(* IEC 61131-3 sources: vespera/src/DUT, 16 files *)

(* ---- ST_BunkerHmi.st ---- *)
(* 8 регистров, адрес = 1100 + (индекс-1)*8 *)
TYPE ST_BunkerHmi :
STRUCT
    wSts      : WORD;   (* +0 маски GVL_Const.BS_* *)
    wAlm      : WORD;   (* +1 GVL_Const.BA_SF *)
    wBypass   : WORD;   (* +2 GVL_Const.BY_DVU *)
    uTDvu     : UINT;   (* +3 с *)
    uTRestart : UINT;   (* +4 с *)
    uRes5     : UINT;
    uRes6     : UINT;
    uRes7     : UINT;
END_STRUCT
END_TYPE

(* ---- ST_BunkerIn.st ---- *)
TYPE ST_BunkerIn :
STRUCT
    xDVU : BOOL;   (* 1 = верхний уровень *)
    xDNU : BOOL;   (* 1 = продукт на нижнем уровне (для бункера поз.27 - второй датчик) *)
    xSF  : BOOL;   (* станции TORBA: 1 = автомат пульта управления включен *)
END_STRUCT
END_TYPE

(* ---- ST_BunkerPar.st ---- *)
TYPE ST_BunkerPar :
STRUCT
    wBypass   : WORD;   (* GVL_Const.BY_DVU - ДВУ отключен *)
    uTDvu     : UINT;   (* задержка срабатывания ДВУ, с *)
    uTRestart : UINT;   (* задержка повторного пуска после снятия ДВУ, с *)
END_STRUCT
END_TYPE

(* ---- ST_GlobHmi.st ---- *)
(* Общий блок, %MW0..%MW31 *)
TYPE ST_GlobHmi :
STRUCT
    wCmd        : WORD;  (* +0  маски GVL_Const.G_* *)
    wSts        : WORD;  (* +1  маски GVL_Const.GS_* *)
    wAlm        : WORD;  (* +2  аварийные стопы 1..10 (биты 0..9), 10 пожар, 11 фазы *)
    wWarn       : WORD;  (* +3  маски GVL_Const.GW_* *)
    uHeartbeat  : UINT;  (* +4  счётчик секунд, контроль связи *)
    uTPreStart  : UINT;  (* +5  предпусковой сигнал, с *)
    uTDksGrace  : UINT;  (* +6  разгон до контроля ДКС, с *)
    uTDksPulse  : UINT;  (* +7  нет импульсов ДКС, 0.1 с *)
    uTFcFb      : UINT;  (* +8  нет сигнала работы ПЧ, с *)
    uTFsStart   : UINT;  (* +9  нет статуса фотосепаратора после пуска, с *)
    uTGateMove  : UINT;  (* +10 контроль хода заслонки поз.1, с *)
    uSirenOn    : UINT;  (* +11 1 = аварийная сирена разрешена *)
    uRes        : ARRAY[12..31] OF UINT;
END_STRUCT
END_TYPE

(* ---- ST_GlobPar.st ---- *)
TYPE ST_GlobPar :
STRUCT
    uTPreStart : UINT;
    uTDksGrace : UINT;
    uTDksPulse : UINT;   (* 0.1 с *)
    uTFcFb     : UINT;
    uTFsStart  : UINT;
    uTGateMove : UINT;
    uSirenOn   : UINT;
END_STRUCT
END_TYPE

(* ---- ST_Link.st ---- *)
(* Связь "механизм подаёт на ..." для блокировок и последовательностей *)
TYPE ST_Link :
STRUCT
    iFrom    : INT;    (* индекс механизма-источника *)
    eTo      : INT;    (* GVL_Const.LT_MECH / LT_BUNKER / LT_INVALID *)
    iTo      : INT;    (* индекс механизма или бункера *)
    xProduct : BOOL;   (* TRUE - поток продукта (пауза по ДВУ распространяется назад),
                          FALSE - вспомогательная связь (аспирация, отходы) *)
END_STRUCT
END_TYPE

(* ---- ST_MechCfg.st ---- *)
(* Постоянная конфигурация механизма *)
TYPE ST_MechCfg :
STRUCT
    eKind     : INT;     (* GVL_Const.K_DOL / K_FC / K_GATE / K_FS *)
    xHasQF    : BOOL;    (* контроль автомата защиты (QF/SF) *)
    eDks      : INT;     (* GVL_Const.DKS_NONE / DKS_PULSE / DKS_LEVEL *)
    xHasDSL   : BOOL;    (* датчики сбегания ленты 1 и 2 *)
    xHasDP    : BOOL;    (* датчик подпора *)
    xHasLocal : BOOL;    (* пост местного управления: ключ Авт/Ручн, Пуск, Стоп *)
    xHasEStop : BOOL;    (* аварийный/концевой стоп у механизма *)
    uDefTOn   : UINT;    (* задержка пуска по умолчанию, с *)
    uDefTOff  : UINT;    (* задержка останова по умолчанию, с *)
END_STRUCT
END_TYPE

(* ---- ST_MechHmi.st ---- *)
(* Обмен с панелью по механизму: 16 регистров %MW (только 16-битные поля).
   Адрес = 200 + (индекс-1)*16 + смещение. *)
TYPE ST_MechHmi :
STRUCT
    wCmd           : WORD;  (* +0  команды панели, маски GVL_Const.C_* *)
    wSts           : WORD;  (* +1  состояние, маски GVL_Const.S_* *)
    wAlm           : WORD;  (* +2  аварии (с фиксацией), маски GVL_Const.A_* *)
    wBypass        : WORD;  (* +3  отключение датчиков (запись с паролем) *)
    uTOn           : UINT;  (* +4  задержка пуска, с *)
    uTOff          : UINT;  (* +5  задержка останова, с *)
    uToInterval    : UINT;  (* +6  интервал ТО, ч *)
    uHoursSinceTO  : UINT;  (* +7  наработка после ТО, ч *)
    uHoursTotal    : UINT;  (* +8  наработка всего, ч *)
    uMinutes       : UINT;  (* +9  минуты наработки (0..59) *)
    iState         : INT;   (* +10 0 стоп, 1 пуск, 2 работа, 3 останов, 4 авария, 5 местное *)
    uRes11         : UINT;
    uRes12         : UINT;
    uRes13         : UINT;
    uRes14         : UINT;
    uRes15         : UINT;
END_STRUCT
END_TYPE

(* ---- ST_MechIn.st ---- *)
(* Логические входы механизма (после учёта полярности в PRG_Inputs) *)
TYPE ST_MechIn :
STRUCT
    xQF       : BOOL;    (* 1 = автомат включен *)
    xDKS      : BOOL;    (* импульсы/уровень датчика контроля скорости *)
    xDSL1     : BOOL;    (* 1 = лента в норме *)
    xDSL2     : BOOL;
    xDP       : BOOL;    (* 1 = подпора нет *)
    xLocal    : BOOL;    (* 1 = ключ поста в положении "ручн." (местное управление) *)
    xLocStart : BOOL;    (* кнопка "Пуск" поста, НО *)
    xLocStop  : BOOL;    (* 1 = кнопка "Стоп" поста не нажата (НЗ) *)
    xEStop    : BOOL;    (* 1 = аварийный/концевой стоп не нажат (НЗ) *)
    xFcFault  : BOOL;    (* 1 = авария ПЧ *)
    xFcReady  : BOOL;    (* 1 = готовность/работа ПЧ *)
    xFb1      : BOOL;    (* заслонка: открыта;  фотосепаратор: статус "работа" *)
    xFb2      : BOOL;    (* заслонка: закрыта;  фотосепаратор: внешнее управление *)
    xErr      : BOOL;    (* фотосепаратор: критическая ошибка *)
    xLocOpen  : BOOL;    (* заслонка: кнопка "Открыть" поста *)
    xLocClose : BOOL;    (* заслонка: кнопка "Закрыть" поста *)
    xAux      : BOOL;    (* фотосепаратор: компрессор в работе (автомат включен) *)
END_STRUCT
END_TYPE

(* ---- ST_MechOut.st ---- *)
TYPE ST_MechOut :
STRUCT
    qRun    : BOOL;      (* пуск двигателя / пуск ПЧ *)
    qPower  : BOOL;      (* включить питание ПЧ (сетевой контактор) *)
    qReset  : BOOL;      (* сброс аварии ПЧ, импульс *)
    qOpen   : BOOL;      (* заслонка: открыть *)
    qClose  : BOOL;      (* заслонка: закрыть *)
    qOn     : BOOL;      (* фотосепаратор: импульс "Включить" *)
    qOff    : BOOL;      (* фотосепаратор: импульс "Выключить" *)
    qEnable : BOOL;      (* фотосепаратор: разрешить секции 1-3 *)
END_STRUCT
END_TYPE

(* ---- ST_MechPar.st ---- *)
(* Уставки и счётчики механизма, хранятся в RETAIN *)
TYPE ST_MechPar :
STRUCT
    uTOn         : UINT;     (* задержка пуска, с *)
    uTOff        : UINT;     (* задержка останова, с *)
    uToInterval  : UINT;     (* интервал ТО, ч; 0 = не контролировать *)
    wBypass      : WORD;     (* отключенные датчики, маски GVL_Const.BY_* *)
    udSecTotal   : UDINT;    (* наработка всего, с *)
    udSecSinceTO : UDINT;    (* наработка после ТО, с *)
END_STRUCT
END_TYPE

(* ---- ST_RouteHmi.st ---- *)
(* 4 регистра, адрес = 100 + (номер-1)*4 *)
TYPE ST_RouteHmi :
STRUCT
    wCmd      : WORD;  (* +0 маски GVL_Const.RC_* *)
    wSts      : WORD;  (* +1 маски GVL_Const.RS_* *)
    iNotReady : INT;   (* +2 причина отказа в пуске: 1..37 механизм, 101..105 клапан, 201..207 бункер,
                          -1 общая авария/цепь управления, -2 конфликт маршрутов, -3 ошибка конфигурации *)
    iState    : INT;   (* +3 0 стоп, 1 предпусковой сигнал, 2 перевод клапанов, 3 работа, 4 останов *)
END_STRUCT
END_TYPE

(* ---- ST_ValveHmi.st ---- *)
(* 8 регистров, адрес = 1000 + (индекс-1)*8 *)
TYPE ST_ValveHmi :
STRUCT
    wCmd   : WORD;   (* +0 маски GVL_Const.VC_* *)
    wSts   : WORD;   (* +1 маски GVL_Const.VS_* *)
    wAlm   : WORD;   (* +2 маски GVL_Const.VA_* *)
    uTMove : UINT;   (* +3 контроль времени перевода, с *)
    uRes4  : UINT;
    uRes5  : UINT;
    uRes6  : UINT;
    uRes7  : UINT;
END_STRUCT
END_TYPE

(* ---- ST_ValveIn.st ---- *)
TYPE ST_ValveIn :
STRUCT
    xSF : BOOL;  (* 1 = автомат привода включен *)
    xS1 : BOOL;  (* датчик положения 1 *)
    xS2 : BOOL;  (* датчик положения 2 *)
END_STRUCT
END_TYPE

(* ---- ST_ValveOut.st ---- *)
TYPE ST_ValveOut :
STRUCT
    q1 : BOOL;   (* перевод в положение 1 *)
    q2 : BOOL;   (* перевод в положение 2 *)
END_STRUCT
END_TYPE

(* ---- ST_ValvePar.st ---- *)
TYPE ST_ValvePar :
STRUCT
    uTMove : UINT;   (* контроль времени перевода, с *)
END_STRUCT
END_TYPE
